(* IEC 61131-3 sources: STAR-PLC-Agent/results/raw/local_validation_20261110/SELF001_mutant/compile, 1 file *)

(* ---- FB_Task.st ---- *)
FUNCTION_BLOCK FB_Task
VAR_INPUT
    Start : BOOL;
    Stop : BOOL;
    GuardClosed : BOOL;
END_VAR
VAR_OUTPUT
    Run : BOOL := FALSE;
END_VAR

Run := FALSE;
END_FUNCTION_BLOCK
